// TIA Portal V20 export
TYPE "Ablauf Positionen"
   STRUCT
      Position_Ein_Aus : Bool;   // Position Ein Aus
      Freigabe_Position : Bool;   // Freigabe Position
      Fertigmeldung_Position : Bool;   // Fertigmeldung Position
      Station_in_Grundstellung : Bool;   // Station in Grundstellung
      INIT_Ablauf_Station : Bool;   // Graph7 Schrittkette wird bei VKE=1 zurückgesetzt
      Schrittkette_aktiv : Bool;   // Bit wird im Initialschritt oder bei Richten 0 und im Ersten Schritt VKE=1
      Richten_nach_Not_Aus : Bool;   // Bit wird gesetzt wenn Not-Aus aktiv und Rückgesetzt über Richtenablauf
      Frei : Bool;
      Messung_GUT_POS : Bool;   // Messung GUT-ausgewertet auf Position
      Messung_SCHLECHT_1_POS : Bool;   // Messung Schlecht-ausgewertet auf Position
      Messung_SCHLECHT_2_POS : Bool;   // Messung Schlecht-ausgewertet auf Position
      Schrittnummer : Int;   // Schrittnummer der Ablaufkeitte im Graph7
      Schrittkettenmerker : Array[0..15] of Bool;
      Bool1 : Array[0..7] of Bool;
      Byte1 : Array[0..7] of Byte;
      Anzahl_Messungen_IST : Int;   // Wiederholungshäufigkeit IST der Messung
      Anzahl_Messungen_SOLL : Int;   // Wiederholungshäufigkeit SOLL der Messungen
      INT2 : Array[0..7] of Int;
      Realwert1 : Real;   // Realwert 1
      Realwert2 : Real;   // Realwert 2
      Realwert3 : Real;   // Realwert 3
      Realwert4 : Real;   // Realwert 4
   END_STRUCT;
END_TYPE
